// Mitsubishi GX Works2 project: Section 3 Circuit   PLC: FX3G

PROGRAM MAIN
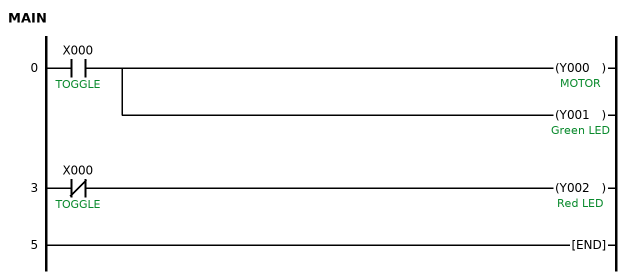
0     LD      X000  ; TOGGLE
      OUT     Y000  ; MOTOR
      OUT     Y001  ; Green LED
3     LDI     X000  ; TOGGLE
      OUT     Y002  ; Red LED
5     END
END_PROGRAM
